Fanuc KAREL source: ka00155.KL

-- PROVISIONAL review KL for V1013-1; original PC SHA256 4288bb402085dc14ce8ff8f7878c6f5aba4d466643ab461e8a74d2e0d729899d
-- Incomplete behavior may be omitted. Consult companion uncertainty JSON. Do not deploy.
PROGRAM KA00155
%NOLOCKGROUP
-- UNRESOLVED_DECL SRC type=002011
-- UNRESOLVED_DECL DST type=002011
BEGIN
  -- UNRESOLVED_PC offsets 5-19; opcodes 22,22,1E
  -- UNRESOLVED_PC offsets 24-28; opcodes 7F
END KA00155
